// TIA Portal V21 export
// export: Created 2026-11-10T19:11:37.2774401Z, ExportSetting WithDefaults, DisplayName Totally Integrated Automation Portal, DisplayVersion V21 Update 3, DisplayName STEP 7 Professional, DisplayVersion V21 Update 3, DisplayName STEP 7 Safety, DisplayVersion V21, DisplayName Tech WebApplication, DisplayVersion V21, DisplayName WinCC Basic/Comfort/Advanced, DisplayVersion V21 Update 3, DisplayName WinCC Unified, DisplayVersion V21 Update 3
DATA_BLOCK "DB_DCAT"   // DB23
// stored: AutoNumber true, DBAccessibleFromOPCUA true, DBAccessibleFromWebserver true, InstanceOfName DCAT, OfSystemLibElement DCAT, OfSystemLibVersion 2.1
"DCAT"
   // VAR_INPUT
   //    CMD : Bool;
   //    O_FB : Bool;
   //    C_FB : Bool;
   // END_VAR
   // VAR_OUTPUT
   //    Q : Bool;
   //    OA : Bool;
   //    CA : Bool;
   // END_VAR
   // VAR
   //    ET : DInt;
   //    PT : DInt;
   //    PREV_TIME : DWord;
   //    CMD_HIS : Bool;
   // END_VAR
BEGIN
END_DATA_BLOCK
